(* IEC 61131-3 sources: volt/packages/volt-lsp-iec/test-corpus/pro2193/Device/Plc Logic/Application/09 Misc/Library Manager/TCP, 10 files *)

(* ---- ERROR.dut ---- *)
TYPE ERROR :
(
	NO_ERROR,
	TIME_OUT,
	PENDING,
	INVALID_HANDLE,
	INVALID_IPADDRESS,
	CONNECT_FAILED,
	HOST_NOT_FOUND,
	TCP_OPEN_ERROR,
	NO_STREAMS_TO_LISTEN,
	ADDR_NOT_AVAILABLE,
	CONNECTION_LOST,
	STREAM_STATE_ERROR,
	GET_OPTION_FAILED,
	SET_OPTION_FAILED,
	IOCTL_FAILED,
	RECEIVE_ERROR,
	SEND_ERROR,
	FD_SET_INIT_FAILED
);
END_TYPE

(* ---- SOCKADDR.dut ---- *)
TYPE SOCKADDR :
STRUCT
	SIN_FAMILY : INT;
	SIN_PORT : UINT;
	SIN_ADDR : UDINT;
	SIN_ZERO : ARRAY [0..7] OF BYTE;
END_STRUCT
END_TYPE

(* ---- STREAM_STATE.dut ---- *)
TYPE STREAM_STATE :
(
	CLOSED := 0,
	CONNECTING,
	LISTENING,
	OPEN,
	FAILED
);
END_TYPE

(* ---- CONSTANTS.gvl ---- *)
VAR_GLOBAL
	GC_DIBACKLOG : DINT := 64;
END_VAR

(* ---- VARIABLES.gvl ---- *)
VAR_GLOBAL
	G_BERRORREUSEPORTGIVEN : BOOL := FALSE;
END_VAR

(* ---- UDINT_TO_IPSTRING.pou ---- *)
FUNCTION UDINT_TO_IPSTRING : STRING
VAR_INPUT
	UDIIPADDRESS : UDINT;
END_VAR
END_FUNCTION

(* ---- CONNECTOR.pou ---- *)
FUNCTION_BLOCK CONNECTOR
VAR
	_HSOCKET : SysTypes.RTS_IEC_HANDLE := SysTypes.RTS_INVALID_HANDLE;
	_UDICLIENTIPADDRESS : UDINT;
	_STREAM : Stream;
	_UDIIPADDRESS : UDINT;
	_UIPORT : UINT;
	_XINITIALIZED : BOOL;
	_XCONNECTED : BOOL;
	_XOPEN : BOOL;
	IPADDRESS : STRING;
	PORT : UINT;
END_VAR
END_FUNCTION_BLOCK

METHOD CONNECT : ERROR
VAR_INPUT
	SIPADDRESS : STRING;
	UIPORT : UINT;
END_VAR
VAR_OUTPUT
	PSTREAM : POINTER TO Stream;
END_VAR
END_METHOD

METHOD DISCONNECT : ERROR
END_METHOD

METHOD FB_EXIT : BOOL
VAR_INPUT
	BINCOPYCODE : BOOL;
END_VAR
END_METHOD

METHOD INITIALIZESOCKET : ERROR
VAR_INPUT
	SIPADDRESS : STRING;
	UIPORT : UINT;
END_VAR
END_METHOD

METHOD RESET
END_METHOD

METHOD RESOLVEHOSTNAME : ERROR
VAR_INPUT
	SHOSTNAME : STRING;
END_VAR
VAR_OUTPUT
	SIPADDRESS : STRING;
END_VAR
END_METHOD

METHOD SETADAPTER : ERROR
VAR_INPUT
	SIPADDRESS : STRING;
END_VAR
END_METHOD

(* ---- LISTENER.pou ---- *)
FUNCTION_BLOCK LISTENER
VAR
	_HLISTENSOCKET : SysTypes.RTS_IEC_HANDLE := SysTypes.RTS_INVALID_HANDLE;
	_LISTENFD_SET : SysSocket.SOCKET_FD_SET;
	_UIPORT : UINT;
	_UDIIPADDRESS : UDINT;
	_XSTARTED : BOOL;
	_XLISTENING : BOOL;
	IPADDRESS : STRING;
	PORT : UINT;
	SOCKET : RTS_IEC_HANDLE;
END_VAR
END_FUNCTION_BLOCK

METHOD ACCEPT : ERROR
VAR_INPUT
	PSTREAM : POINTER TO Stream;
END_VAR
END_METHOD

METHOD FB_EXIT : BOOL
VAR_INPUT
	BINCOPYCODE : BOOL;
END_VAR
END_METHOD

METHOD LISTEN : ERROR
END_METHOD

METHOD START : ERROR
VAR_INPUT
	SIPADDRESS : STRING;
	UIPORT : UINT;
END_VAR
END_METHOD

METHOD STOP : ERROR
END_METHOD

(* ---- SELECT.pou ---- *)
FUNCTION_BLOCK SELECT
END_FUNCTION_BLOCK

METHOD CHECK : ERROR
VAR_INPUT
	ITIMEOUT : INT;
END_VAR
VAR_OUTPUT
	DIREADY : DINT;
END_VAR
VAR_IN_OUT
	STRRECVSET : SysSocket.SOCKET_FD_SET;
	STRSENDSET : SysSocket.SOCKET_FD_SET;
	STRERRORSET : SysSocket.SOCKET_FD_SET;
END_VAR
END_METHOD

METHOD CHECKERROR : ERROR
VAR_INPUT
	ITIMEOUT : INT;
END_VAR
VAR_OUTPUT
	DIREADY : DINT;
END_VAR
VAR_IN_OUT
	SOCKETFD_SET : SysSocket.SOCKET_FD_SET;
END_VAR
END_METHOD

METHOD CHECKRECEIVE : ERROR
VAR_INPUT
	ITIMEOUT : INT;
END_VAR
VAR_OUTPUT
	DIREADY : DINT;
END_VAR
VAR_IN_OUT
	SOCKETFD_SET : SysSocket.SOCKET_FD_SET;
END_VAR
END_METHOD

METHOD CHECKSEND : ERROR
VAR_INPUT
	ITIMEOUT : INT;
END_VAR
VAR_OUTPUT
	DIREADY : DINT;
END_VAR
VAR_IN_OUT
	SOCKETFD_SET : SysSocket.SOCKET_FD_SET;
END_VAR
END_METHOD

(* ---- STREAM.pou ---- *)
FUNCTION_BLOCK STREAM
VAR
	_HSOCKET : SysTypes.RTS_IEC_HANDLE := SysTypes.RTS_INVALID_HANDLE;
	_ESTATE : STREAM_STATE;
	_TCPSELECT : Select;
	_IPADDR : SysSocket.INADDR;
	_PUSHBACK1READBYTE_DATA : BYTE;
	_PUSHBACK1READBYTE_CALLED : BOOL;
	IPADDRESS : SysSocket.INADDR;
	SOCKET : SysTypes.RTS_IEC_HANDLE;
	STATE : STREAM_STATE;
END_VAR
END_FUNCTION_BLOCK

METHOD CHECKCONNECTIVITY : BOOL
END_METHOD

METHOD CHECKRECEIVE : BOOL
END_METHOD

METHOD CHECKSEND : BOOL
END_METHOD

METHOD CLOSE : ERROR
END_METHOD

METHOD CREATE : ERROR
VAR_INPUT
	HSOCKET : SysTypes.RTS_IEC_HANDLE;
END_VAR
END_METHOD

METHOD FB_EXIT : BOOL
VAR_INPUT
	BINCOPYCODE : BOOL;
END_VAR
END_METHOD

METHOD FDISSET : BOOL
VAR_INPUT
	SOCKETFD_SET : SysSocket.SOCKET_FD_SET;
END_VAR
END_METHOD

METHOD FDSET
VAR_IN_OUT
	SOCKETFD_SET : SysSocket.SOCKET_FD_SET;
END_VAR
END_METHOD

METHOD GETOPTION : ERROR
VAR_INPUT
	DIOPTION : DINT;
END_VAR
VAR_OUTPUT
	DIVALUE : DINT;
END_VAR
END_METHOD

METHOD IOCONTROL : ERROR
VAR_INPUT
	DICOMMAND : DINT;
END_VAR
VAR_IN_OUT
	DIPARAMETER : DINT;
END_VAR
END_METHOD

METHOD RECEIVE : ERROR
VAR_INPUT
	PBYBUFFER : POINTER TO BYTE;
	DIBUFFERSIZE : __XINT;
END_VAR
VAR_OUTPUT
	DIRECEIVED : __XINT;
END_VAR
END_METHOD

METHOD RESET
END_METHOD

METHOD SEND : ERROR
VAR_INPUT
	PBYBUFFER : POINTER TO BYTE;
	DIBUFFERSIZE : __XINT;
END_VAR
VAR_OUTPUT
	DISENT : __XINT;
END_VAR
END_METHOD

METHOD SETOPTION : ERROR
VAR_INPUT
	DIOPTION : DINT;
	DIVALUE : DINT;
END_VAR
END_METHOD

METHOD GETPUSHBACK1READBYTE
VAR_OUTPUT
	DATA : BYTE;
	CALLED : BOOL;
END_VAR
END_METHOD

METHOD SETPUSHBACK1READBYTE
VAR_INPUT
	DATA : BYTE;
	CALLED : BOOL;
END_VAR
END_METHOD
